(* Logix 5000 project; controller MECO9497 vendor 1 type 14 code 106 rev 21.11; software revision 21.00; part 2 of 4 *)
(* tags used below, declared in another part *)
   AAH_200 : BOOL;
   AAH_200_DELAY : TIMER;
   AAH_200_SP : REAL;
   ACKNOWLEDGE : BOOL;
   ALARM_ACK_OIT : BOOL;
   ALARM_RESET_OIT : BOOL;
   ALERT_ALARM_SU_DELAY : TIMER;
   AT_200_EU : REAL;
   COMP_AMP_ALRM_DELAY_TMR : TIMER;
   COMPRESSOR_START_CMD : BOOL;
   D_V_REMOTE_START : BOOL;
   DIST_COND_ALRM_STARTUP_TMR : TIMER;
   DSTLT_STORAGE_ENABLE_MAP : BOOL;
   DSTLT_STORAGE_ENABLE_OIT : BOOL;
   DSTLT_TEMP_ALRM_SU_DELAY : TIMER;
   E_Stop : ALIAS FOR Local:1:I.Data.0;
   E_Stop_DI_MAP : BOOL;
   ENGINEER : BOOL;
   EVAP_PRESS_CV_LIMIT : BOOL;
   EVAP_PRESS_CV_PERMISSIVE : REAL;
   EVAP_PRESS_RAMP_ONE_SHOT : BOOL;
   EVAP_PRESS_RAMP_TIMER : TIMER;
   EVAP_PRESSURE_CV_PERM : BOOL;
   EVAP_RAMP_COMPLETE : BOOL;
   EVAP_RAMP_ENABLE_DELAY_TIMER : TIMER;
   FEED_LVL_CV_LIMIT : BOOL;
   FEED_LVL_CV_LIMIT_SHUTDOWN : BOOL;
   FEED_LVL_CV_LIMIT_SHUTDOWN_DELAY : TIMER;
   FEED_LVL_CV_LIMIT_SHUTDOWN_LATCH : BOOL;
   FEED_LVL_ONE_SHOT : BOOL;
   FEED_TEM_SD_LATCH : BOOL;
   FEED_TEM_SD_TIMER : TIMER;
   FEED_TEMP_SD_ONS : BOOL;
   FEED_TEMP_STEP_DELAY : TIMER;
   HOT_STANDBY : BOOL;
   IAL_100 : BOOL;
   IAL_100_CTR : COUNTER;
   IAL_100_DELAY : TIMER;
   IAL_100_SP : REAL;
   INITIAL_SCAN_SYS_RESET : BOOL;
   INITIAL_START_STEAM_LIMIT_TMR : TIMER;
   IY_100_EU : REAL;
   LAAH_100 : BOOL;
   LAAH_100_DELAY : TIMER;
   LAAH_100_SP : DINT;
   LAAL_100 : BOOL;
   LAAL_100_DELAY : TIMER;
   LAAL_100_SP : DINT;
   LAH_100 : BOOL;
   LAH_100_AUX : BOOL;
   LAH_100_DELAY : TIMER;
   LAH_100_SP : REAL;
   LAL_100 : BOOL;
   LAL_100_DELAY : TIMER;
   LAL_100_SP : REAL;
   LB_OIL_LOW_PRESS_ALRM_DELAY : TIMER;
   LCV_100_INTERLOCK : BOOL;
   LIC_100 : PID;
   LIC_1000_CV1 : REAL;
   LIC_100_A_M_OIT : BOOL;
   LIC_100_CV2 : REAL;
   LIC_100_CV_H : BOOL;
   LIC_100_CV_N : BOOL;
   LIC_100_CV_OIT : REAL;
   LIC_100_FINAL_SP : REAL;
   LIC_100_FINAL_SP_EU : REAL;
   LIC_100_GAIN_H : BOOL;
   LIC_100_GAIN_N : BOOL;
   LIC_100_GAIN_OIT : REAL;
   LIC_100_RATE_H : BOOL;
   LIC_100_RATE_N : BOOL;
   LIC_100_RATE_OIT : REAL;
   LIC_100_RESET_H : BOOL;
   LIC_100_RESET_N : BOOL;
   LIC_100_RESET_OIT : REAL;
   LIC_100_SP_CONV : REAL;
   LIC_100_SP_EU : REAL;
   LIC_100_SP_H : BOOL;
   LIC_100_SP_N : BOOL;
   LIC_100_SP_OIT : REAL;
   LIC_100_STBY_SP : REAL;
   LIC_100_STBY_SP_EU : REAL;
   LIC_100_STBY_SP_H : BOOL;
   LIC_100_STBY_SP_N : BOOL;
   LIC_100_STBY_SP_OIT : REAL;
   LT_100_AI : ALIAS FOR Local:3:I.Ch3Data;
   LT_100_EU : REAL;
   LT_100_EU_SPAN : REAL;
   LT_100_EU_ZERO : REAL;
   M1_DI : ALIAS FOR Local:1:I.Data.1;
   M1_DI_MAP : BOOL;
   M2_DI : ALIAS FOR Local:1:I.Data.2;
   M2_DI_MAP : BOOL;
   M4_DI : ALIAS FOR Local:1:I.Data.4;
   M4_DI_MAP : BOOL;
   MAINTENANCE : BOOL;
   MCB : BOOL;
   OP_SWTCH_AUTO_DI : ALIAS FOR Local:1:I.Data.14;
   OP_SWTCH_AUTO_DI_MAP : BOOL;
   OP_SWTCH_MANUAL_DI : ALIAS FOR Local:1:I.Data.13;
   OP_SWTCH_MANUAL_DI_MAP : BOOL;
   OPERATOR : BOOL;
   PAAH_103 : BOOL;
   PAAH_103_DELAY : TIMER;
   PAAH_103_SP : REAL;
   PAAL_103 : BOOL;
   PAAL_103_DELAY : TIMER;
   PAAL_103_SP : REAL;
   PAH_103 : BOOL;
   PAH_103_AUX : BOOL;
   PAH_103_DELAY : TIMER;
   PAH_103_SP : REAL;
   PAL_103 : BOOL;
   PAL_103_DELAY : TIMER;
   PAL_103_SP : REAL;
   PAL_700 : BOOL;
   PAL_700_ALRM_DELAY : TIMER;
   PCV_103_INTERLOCK : BOOL;
   PIC_103 : PID;
   PIC_103_A_M_OIT : BOOL;
   PIC_103_CV_H : BOOL;
   PIC_103_CV_N : BOOL;
   PIC_103_CV_OIT : REAL;
   PIC_103_FINAL_SP : REAL;
   PIC_103_GAIN_H : BOOL;
   PIC_103_GAIN_N : BOOL;
   PIC_103_GAIN_OIT : REAL;
   PIC_103_RATE_H : BOOL;
   PIC_103_RATE_N : BOOL;
   PIC_103_RATE_OIT : REAL;
   PIC_103_RESET_H : BOOL;
   PIC_103_RESET_N : BOOL;
   PIC_103_RESET_OIT : REAL;
   PIC_103_SP_CONV : REAL;
   PIC_103_SP_EU : REAL;
   PIC_103_SP_H : BOOL;
   PIC_103_SP_N : BOOL;
   PIC_103_SP_OIT : REAL;
   PIC_103_STBY_SP : REAL;
   PIC_103_STBY_SP_EU : REAL;
   PIC_103_STBY_SP_H : BOOL;
   PIC_103_STBY_SP_N : BOOL;
   PIC_103_STBY_SP_OIT : REAL;
   PSL_700_DI : ALIAS FOR Local:1:I.Data.7;
   PT_103_AI : ALIAS FOR Local:3:I.Ch0Data;
   PT_103_EU : REAL;
   PT_103_EU_SPAN : REAL;
   PT_103_EU_ZERO : REAL;
   PT_103_HIGH : REAL;
   RESET : BOOL;
   SECURITY_ENABLED : BOOL;
   TAH_700 : BOOL;
   TAH_700_ALRM_DELAY : TIMER;
   TAL_200 : BOOL;
   TAL_200_DELAY : TIMER;
   TAL_200_SP : REAL;
   TIC_102 : PID;
   TIC_102_A_M_OIT : BOOL;
   TIC_102_CV_H : BOOL;
   TIC_102_CV_MIN_LIMIT : BOOL;
   TIC_102_CV_N : BOOL;
   TIC_102_CV_OIT : REAL;
   TIC_102_CV_SU_REM : DINT;
   TIC_102_CV_SU_TIMER : TIMER;
   TIC_102_GAIN_H : BOOL;
   TIC_102_GAIN_N : BOOL;
   TIC_102_GAIN_OIT : REAL;
   TIC_102_MINCV1 : REAL;
   TIC_102_MINCV2 : REAL;
   TIC_102_MINCV3 : REAL;
   TIC_102_RATE_H : BOOL;
   TIC_102_RATE_N : BOOL;
   TIC_102_RATE_OIT : REAL;
   TIC_102_RESET_H : BOOL;
   TIC_102_RESET_N : BOOL;
   TIC_102_RESET_OIT : REAL;
   TIC_102_SP_CONV : REAL;
   TIC_102_SP_EU : REAL;
   TIC_102_SP_H : BOOL;
   TIC_102_SP_N : BOOL;
   TIC_102_SP_OIT : REAL;
   TIC_102_START_CV_TIMER_SP_H : BOOL;
   TIC_102_START_CV_TIMER_SP_N : BOOL;
   TIC_102_START_CV_TIMER_SP_O : REAL;
   TSH_700_DI : ALIAS FOR Local:1:I.Data.8;
   TT_102_EU_SPAN : REAL;
   TT_102_EU_ZERO : REAL;
   TT_200_EU : REAL;
   UNIT_REMOTE_START_DI : ALIAS FOR Local:1:I.Data.12;
   UNIT_REMOTE_START_MAP : BOOL;
   UNIT_START_DI : ALIAS FOR Local:1:I.Data.10;
   UNIT_START_DI_MAP : BOOL;
   UNIT_STOP_DI : ALIAS FOR Local:1:I.Data.11;
   UNIT_STOP_DI_MAP : BOOL;
(* MainProgram, continued *)

ROUTINE EVAPORATOR_PRESSURE   (* ladder *)
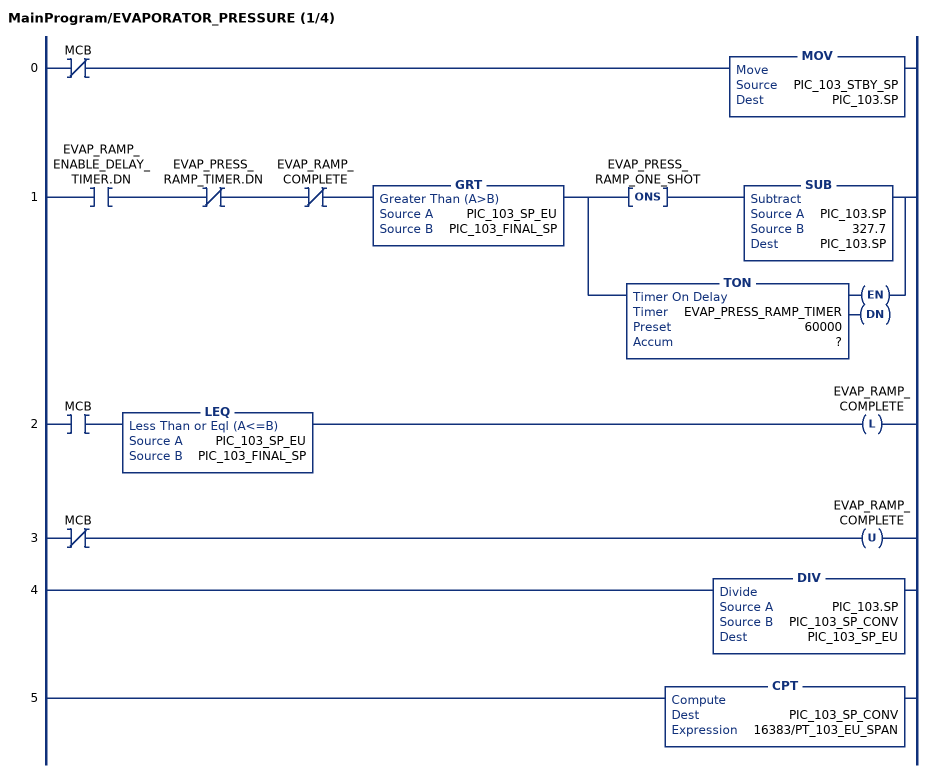
   0: XIO(MCB)MOV(PIC_103_STBY_SP,PIC_103.SP);
   1: XIC(EVAP_RAMP_ENABLE_DELAY_TIMER.DN)XIO(EVAP_PRESS_RAMP_TIMER.DN)XIO(EVAP_RAMP_COMPLETE)GRT(PIC_103_SP_EU,PIC_103_FINAL_SP)[ONS(EVAP_PRESS_RAMP_ONE_SHOT) SUB(PIC_103.SP,327.7,PIC_103.SP) ,TON(EVAP_PRESS_RAMP_TIMER,?,?) ];
   2: XIC(MCB)LEQ(PIC_103_SP_EU,PIC_103_FINAL_SP)OTL(EVAP_RAMP_COMPLETE);
   3: XIO(MCB)OTU(EVAP_RAMP_COMPLETE);
   4: DIV(PIC_103.SP,PIC_103_SP_CONV,PIC_103_SP_EU);
   5: CPT(PIC_103_SP_CONV,16383/PT_103_EU_SPAN);
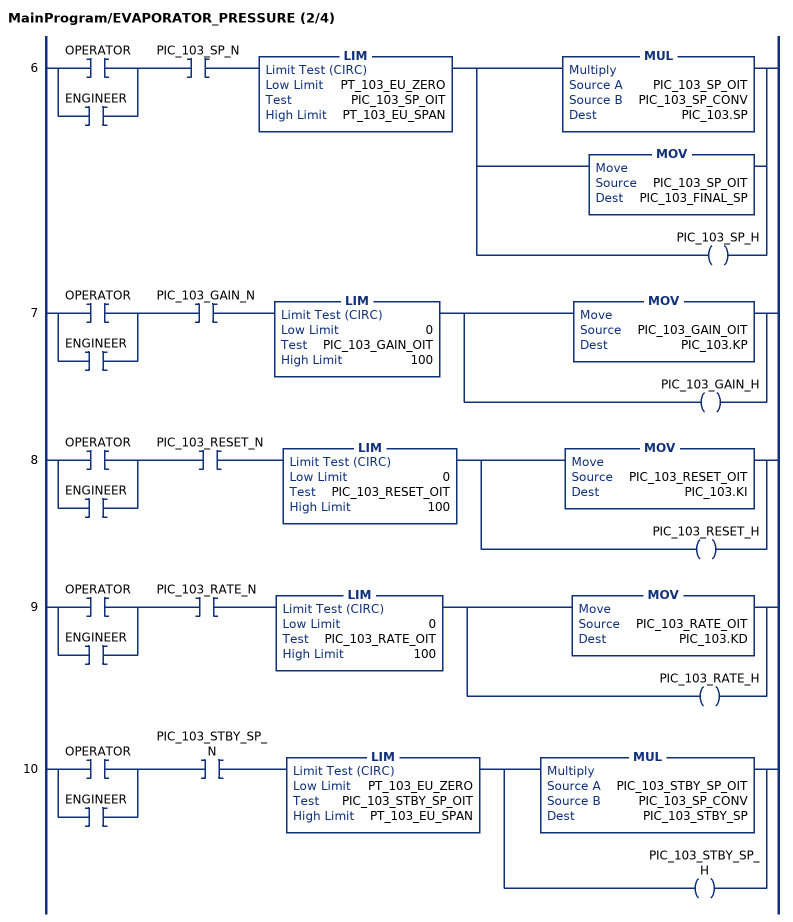
   6: [XIC(OPERATOR) ,XIC(ENGINEER) ]XIC(PIC_103_SP_N)LIM(PT_103_EU_ZERO,PIC_103_SP_OIT,PT_103_EU_SPAN)[MUL(PIC_103_SP_OIT,PIC_103_SP_CONV,PIC_103.SP) ,MOV(PIC_103_SP_OIT,PIC_103_FINAL_SP) ,OTE(PIC_103_SP_H) ];
   7: [XIC(OPERATOR) ,XIC(ENGINEER) ]XIC(PIC_103_GAIN_N)LIM(0,PIC_103_GAIN_OIT,100)[MOV(PIC_103_GAIN_OIT,PIC_103.KP) ,OTE(PIC_103_GAIN_H) ];
   8: [XIC(OPERATOR) ,XIC(ENGINEER) ]XIC(PIC_103_RESET_N)LIM(0,PIC_103_RESET_OIT,100)[MOV(PIC_103_RESET_OIT,PIC_103.KI) ,OTE(PIC_103_RESET_H) ];
   9: [XIC(OPERATOR) ,XIC(ENGINEER) ]XIC(PIC_103_RATE_N)LIM(0,PIC_103_RATE_OIT,100)[MOV(PIC_103_RATE_OIT,PIC_103.KD) ,OTE(PIC_103_RATE_H) ];
   10: [XIC(OPERATOR) ,XIC(ENGINEER) ]XIC(PIC_103_STBY_SP_N)LIM(PT_103_EU_ZERO,PIC_103_STBY_SP_OIT,PT_103_EU_SPAN)[MUL(PIC_103_STBY_SP_OIT,PIC_103_SP_CONV,PIC_103_STBY_SP) ,OTE(PIC_103_STBY_SP_H) ];
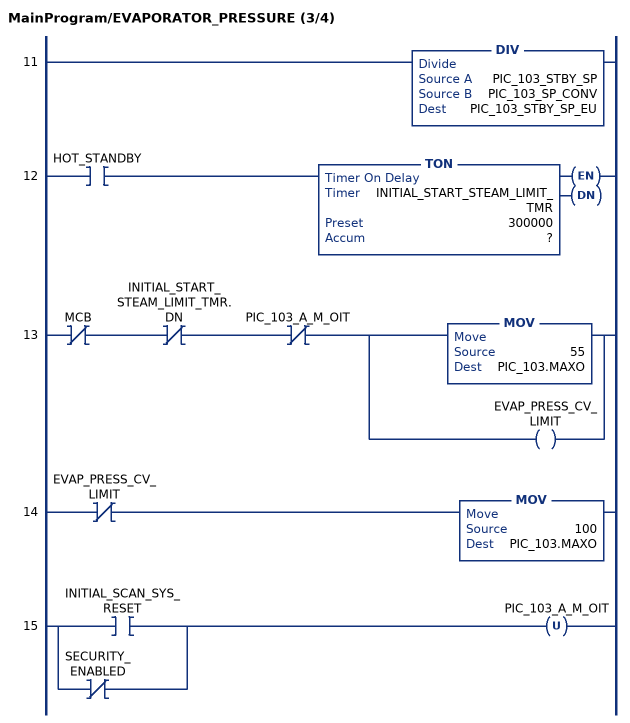
   11: DIV(PIC_103_STBY_SP,PIC_103_SP_CONV,PIC_103_STBY_SP_EU);
   12: XIC(HOT_STANDBY)TON(INITIAL_START_STEAM_LIMIT_TMR,?,?);
   13: XIO(MCB)XIO(INITIAL_START_STEAM_LIMIT_TMR.DN)XIO(PIC_103_A_M_OIT)[MOV(55,PIC_103.MAXO) ,OTE(EVAP_PRESS_CV_LIMIT) ];
   14: XIO(EVAP_PRESS_CV_LIMIT)MOV(100,PIC_103.MAXO);
   15: [XIC(INITIAL_SCAN_SYS_RESET) ,XIO(SECURITY_ENABLED) ]OTU(PIC_103_A_M_OIT);
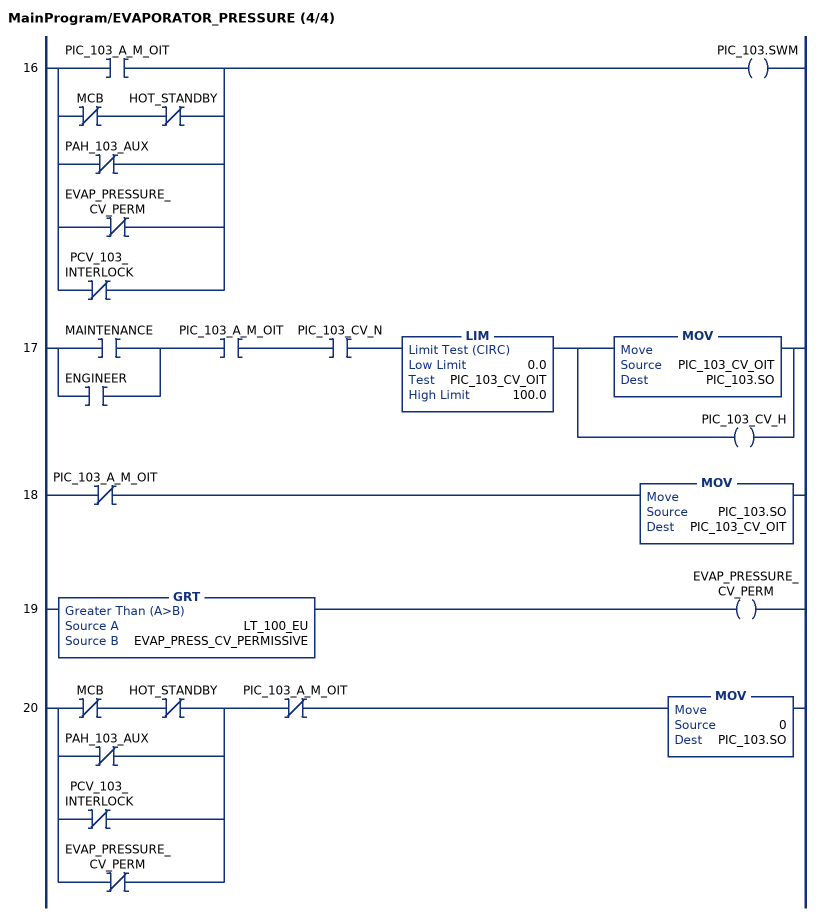
   16: [XIC(PIC_103_A_M_OIT) ,XIO(MCB) XIO(HOT_STANDBY) ,XIO(PAH_103_AUX) ,XIO(EVAP_PRESSURE_CV_PERM) ,XIO(PCV_103_INTERLOCK) ]OTE(PIC_103.SWM);
   17: [XIC(MAINTENANCE) ,XIC(ENGINEER) ]XIC(PIC_103_A_M_OIT)XIC(PIC_103_CV_N)LIM(0.0,PIC_103_CV_OIT,100.0)[MOV(PIC_103_CV_OIT,PIC_103.SO) ,OTE(PIC_103_CV_H) ];
   18: XIO(PIC_103_A_M_OIT)MOV(PIC_103.SO,PIC_103_CV_OIT);
   19: GRT(LT_100_EU,EVAP_PRESS_CV_PERMISSIVE)OTE(EVAP_PRESSURE_CV_PERM);
   20: [XIO(MCB) XIO(HOT_STANDBY) ,XIO(PAH_103_AUX) ,XIO(PCV_103_INTERLOCK) ,XIO(EVAP_PRESSURE_CV_PERM) ]XIO(PIC_103_A_M_OIT)MOV(0,PIC_103.SO);
END_ROUTINE

ROUTINE FEED_LEVEL   (* ladder *)
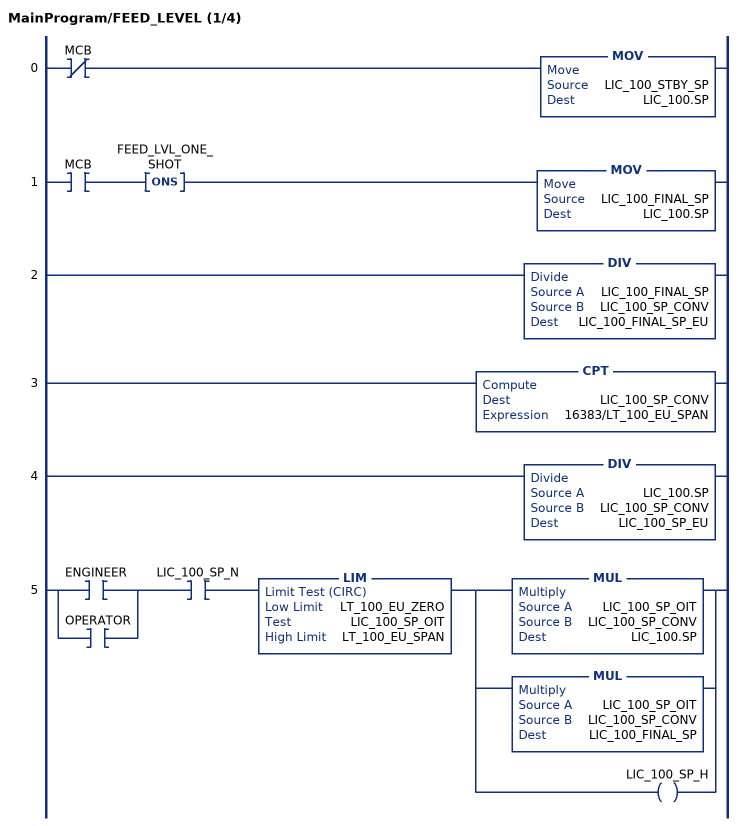
   0: XIO(MCB)MOV(LIC_100_STBY_SP,LIC_100.SP);
   1: XIC(MCB)ONS(FEED_LVL_ONE_SHOT)MOV(LIC_100_FINAL_SP,LIC_100.SP);
   2: DIV(LIC_100_FINAL_SP,LIC_100_SP_CONV,LIC_100_FINAL_SP_EU);
   3: CPT(LIC_100_SP_CONV,16383/LT_100_EU_SPAN);
   4: DIV(LIC_100.SP,LIC_100_SP_CONV,LIC_100_SP_EU);
   5: [XIC(ENGINEER) ,XIC(OPERATOR) ]XIC(LIC_100_SP_N)LIM(LT_100_EU_ZERO,LIC_100_SP_OIT,LT_100_EU_SPAN)[[MUL(LIC_100_SP_OIT,LIC_100_SP_CONV,LIC_100.SP) ,MUL(LIC_100_SP_OIT,LIC_100_SP_CONV,LIC_100_FINAL_SP) ] ,OTE(LIC_100_SP_H) ];
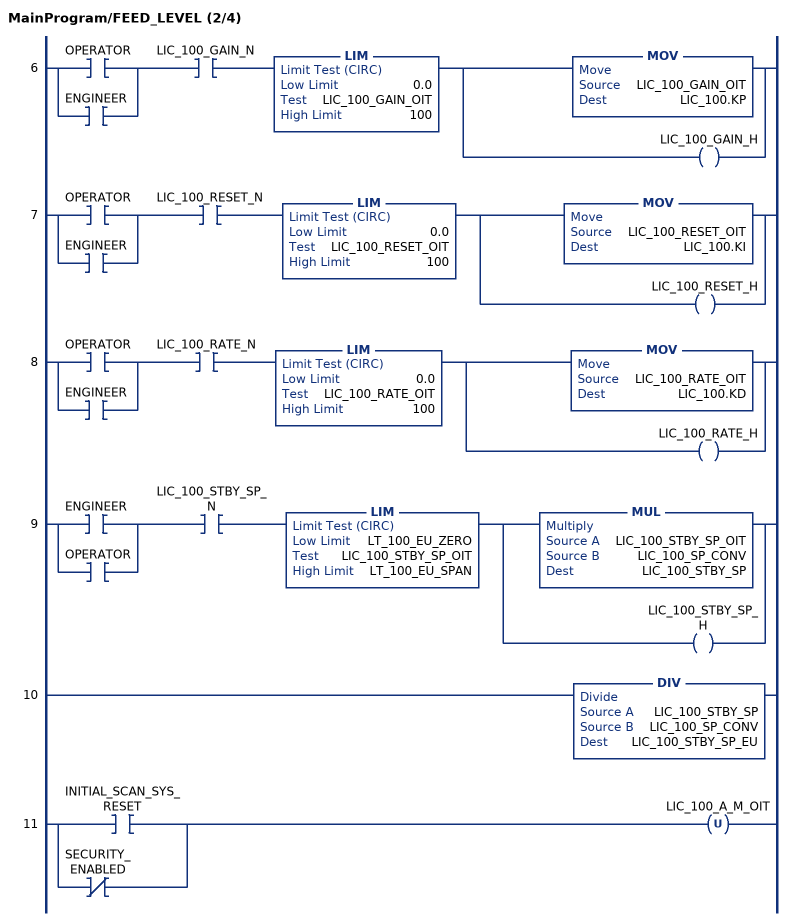
   6: [XIC(OPERATOR) ,XIC(ENGINEER) ]XIC(LIC_100_GAIN_N)LIM(0.0,LIC_100_GAIN_OIT,100)[MOV(LIC_100_GAIN_OIT,LIC_100.KP) ,OTE(LIC_100_GAIN_H) ];
   7: [XIC(OPERATOR) ,XIC(ENGINEER) ]XIC(LIC_100_RESET_N)LIM(0.0,LIC_100_RESET_OIT,100)[MOV(LIC_100_RESET_OIT,LIC_100.KI) ,OTE(LIC_100_RESET_H) ];
   8: [XIC(OPERATOR) ,XIC(ENGINEER) ]XIC(LIC_100_RATE_N)LIM(0.0,LIC_100_RATE_OIT,100)[MOV(LIC_100_RATE_OIT,LIC_100.KD) ,OTE(LIC_100_RATE_H) ];
   9: [XIC(ENGINEER) ,XIC(OPERATOR) ]XIC(LIC_100_STBY_SP_N)LIM(LT_100_EU_ZERO,LIC_100_STBY_SP_OIT,LT_100_EU_SPAN)[MUL(LIC_100_STBY_SP_OIT,LIC_100_SP_CONV,LIC_100_STBY_SP) ,OTE(LIC_100_STBY_SP_H) ];
   10: DIV(LIC_100_STBY_SP,LIC_100_SP_CONV,LIC_100_STBY_SP_EU);
   11: [XIC(INITIAL_SCAN_SYS_RESET) ,XIO(SECURITY_ENABLED) ]OTU(LIC_100_A_M_OIT);
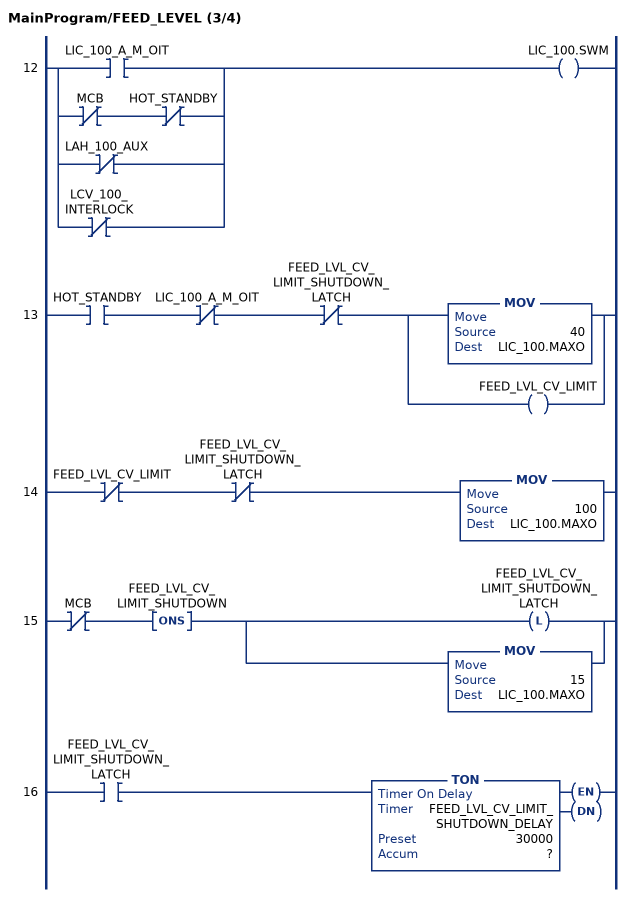
   12: [XIC(LIC_100_A_M_OIT) ,XIO(MCB) XIO(HOT_STANDBY) ,XIO(LAH_100_AUX) ,XIO(LCV_100_INTERLOCK) ]OTE(LIC_100.SWM);
   13: XIC(HOT_STANDBY)XIO(LIC_100_A_M_OIT)XIO(FEED_LVL_CV_LIMIT_SHUTDOWN_LATCH)[MOV(40,LIC_100.MAXO) ,OTE(FEED_LVL_CV_LIMIT) ];
   14: XIO(FEED_LVL_CV_LIMIT)XIO(FEED_LVL_CV_LIMIT_SHUTDOWN_LATCH)MOV(100,LIC_100.MAXO);
   15: XIO(MCB)ONS(FEED_LVL_CV_LIMIT_SHUTDOWN)[OTL(FEED_LVL_CV_LIMIT_SHUTDOWN_LATCH) ,MOV(15,LIC_100.MAXO) ];
   16: XIC(FEED_LVL_CV_LIMIT_SHUTDOWN_LATCH)TON(FEED_LVL_CV_LIMIT_SHUTDOWN_DELAY,?,?);
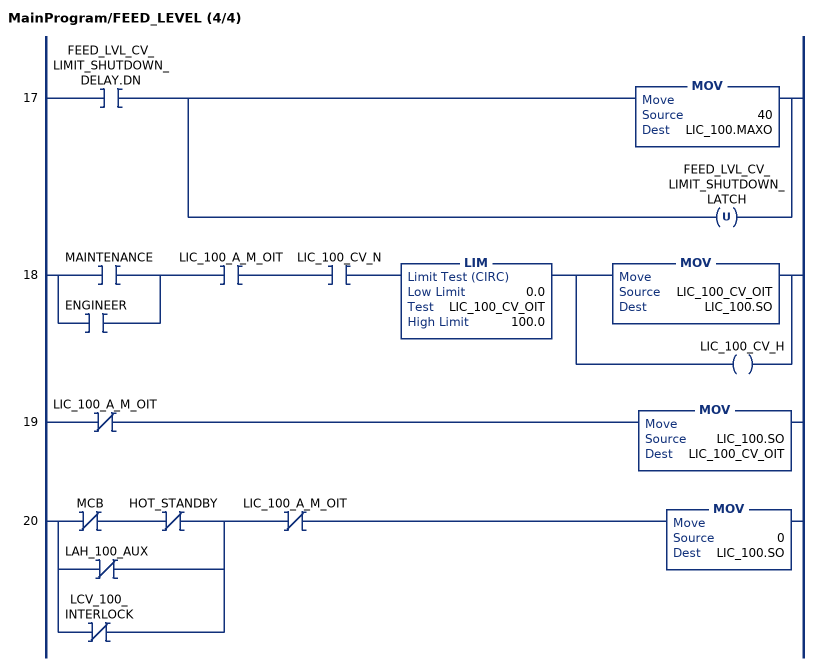
   17: XIC(FEED_LVL_CV_LIMIT_SHUTDOWN_DELAY.DN)[MOV(40,LIC_100.MAXO) ,OTU(FEED_LVL_CV_LIMIT_SHUTDOWN_LATCH) ];
   18: [XIC(MAINTENANCE) ,XIC(ENGINEER) ]XIC(LIC_100_A_M_OIT)XIC(LIC_100_CV_N)LIM(0.0,LIC_100_CV_OIT,100.0)[MOV(LIC_100_CV_OIT,LIC_100.SO) ,OTE(LIC_100_CV_H) ];
   19: XIO(LIC_100_A_M_OIT)MOV(LIC_100.SO,LIC_100_CV_OIT);
   20: [XIO(MCB) XIO(HOT_STANDBY) ,XIO(LAH_100_AUX) ,XIO(LCV_100_INTERLOCK) ]XIO(LIC_100_A_M_OIT)MOV(0,LIC_100.SO);
END_ROUTINE

ROUTINE FEED_TEMPERATURE   (* ladder *)
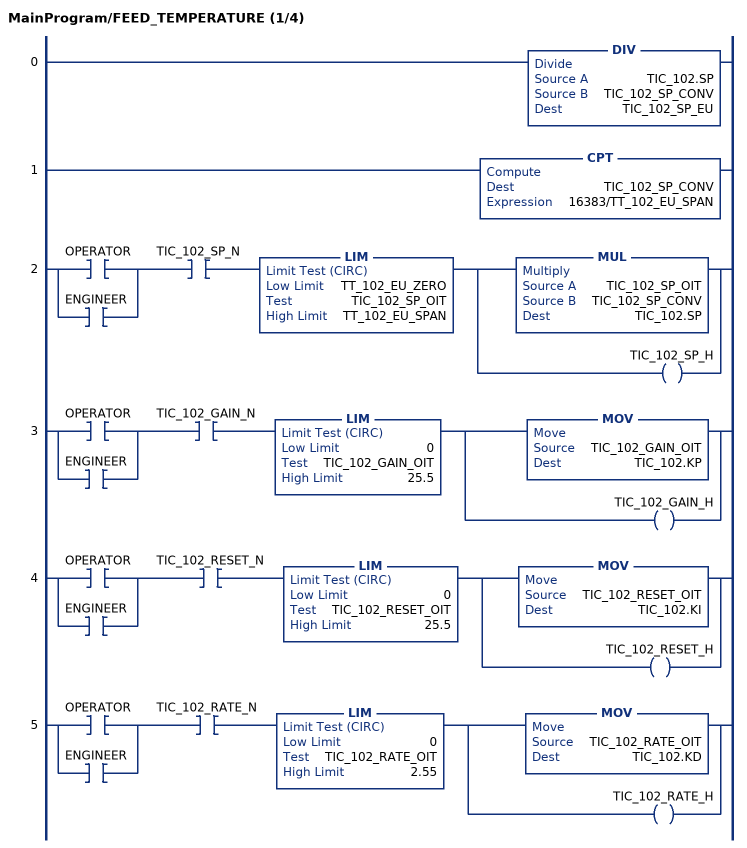
   0: DIV(TIC_102.SP,TIC_102_SP_CONV,TIC_102_SP_EU);
   1: CPT(TIC_102_SP_CONV,16383/TT_102_EU_SPAN);
   2: [XIC(OPERATOR) ,XIC(ENGINEER) ]XIC(TIC_102_SP_N)LIM(TT_102_EU_ZERO,TIC_102_SP_OIT,TT_102_EU_SPAN)[MUL(TIC_102_SP_OIT,TIC_102_SP_CONV,TIC_102.SP) ,OTE(TIC_102_SP_H) ];
   3: [XIC(OPERATOR) ,XIC(ENGINEER) ]XIC(TIC_102_GAIN_N)LIM(0,TIC_102_GAIN_OIT,25.5)[MOV(TIC_102_GAIN_OIT,TIC_102.KP) ,OTE(TIC_102_GAIN_H) ];
   4: [XIC(OPERATOR) ,XIC(ENGINEER) ]XIC(TIC_102_RESET_N)LIM(0,TIC_102_RESET_OIT,25.5)[MOV(TIC_102_RESET_OIT,TIC_102.KI) ,OTE(TIC_102_RESET_H) ];
   5: [XIC(OPERATOR) ,XIC(ENGINEER) ]XIC(TIC_102_RATE_N)LIM(0,TIC_102_RATE_OIT,2.55)[MOV(TIC_102_RATE_OIT,TIC_102.KD) ,OTE(TIC_102_RATE_H) ];
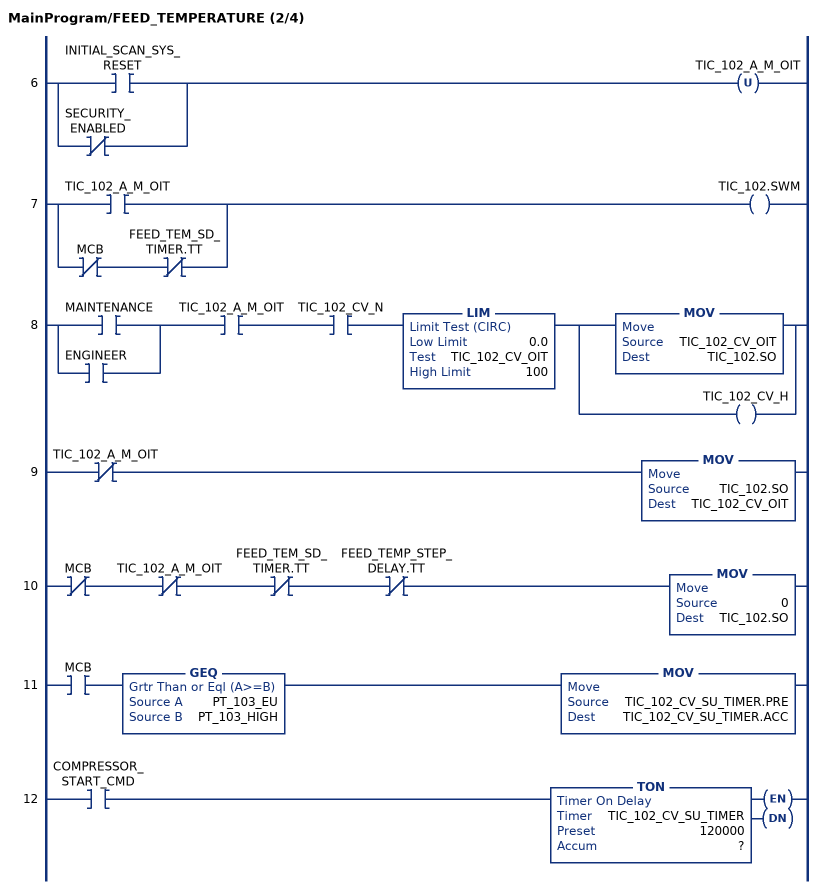
   6: [XIC(INITIAL_SCAN_SYS_RESET) ,XIO(SECURITY_ENABLED) ]OTU(TIC_102_A_M_OIT);
   7: [XIC(TIC_102_A_M_OIT) ,XIO(MCB) XIO(FEED_TEM_SD_TIMER.TT) ]OTE(TIC_102.SWM);
   8: [XIC(MAINTENANCE) ,XIC(ENGINEER) ]XIC(TIC_102_A_M_OIT)XIC(TIC_102_CV_N)LIM(0.0,TIC_102_CV_OIT,100)[MOV(TIC_102_CV_OIT,TIC_102.SO) ,OTE(TIC_102_CV_H) ];
   9: XIO(TIC_102_A_M_OIT)MOV(TIC_102.SO,TIC_102_CV_OIT);
   10: XIO(MCB)XIO(TIC_102_A_M_OIT)XIO(FEED_TEM_SD_TIMER.TT)XIO(FEED_TEMP_STEP_DELAY.TT)MOV(0,TIC_102.SO);
   11: XIC(MCB)GEQ(PT_103_EU,PT_103_HIGH)MOV(TIC_102_CV_SU_TIMER.PRE,TIC_102_CV_SU_TIMER.ACC);
   12: XIC(COMPRESSOR_START_CMD)TON(TIC_102_CV_SU_TIMER,?,?);
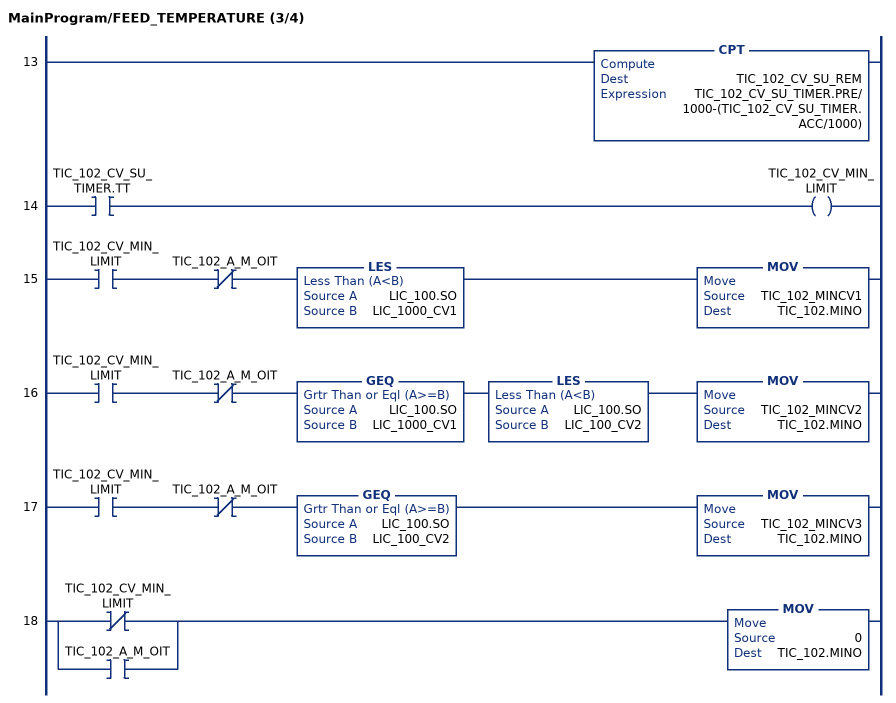
   13: CPT(TIC_102_CV_SU_REM,TIC_102_CV_SU_TIMER.PRE/1000-(TIC_102_CV_SU_TIMER.ACC/1000));
   14: XIC(TIC_102_CV_SU_TIMER.TT)OTE(TIC_102_CV_MIN_LIMIT);
   15: XIC(TIC_102_CV_MIN_LIMIT)XIO(TIC_102_A_M_OIT)LES(LIC_100.SO,LIC_1000_CV1)MOV(TIC_102_MINCV1,TIC_102.MINO);
   16: XIC(TIC_102_CV_MIN_LIMIT)XIO(TIC_102_A_M_OIT)GEQ(LIC_100.SO,LIC_1000_CV1)LES(LIC_100.SO,LIC_100_CV2)MOV(TIC_102_MINCV2,TIC_102.MINO);
   17: XIC(TIC_102_CV_MIN_LIMIT)XIO(TIC_102_A_M_OIT)GEQ(LIC_100.SO,LIC_100_CV2)MOV(TIC_102_MINCV3,TIC_102.MINO);
   18: [XIO(TIC_102_CV_MIN_LIMIT) ,XIC(TIC_102_A_M_OIT) ]MOV(0,TIC_102.MINO);
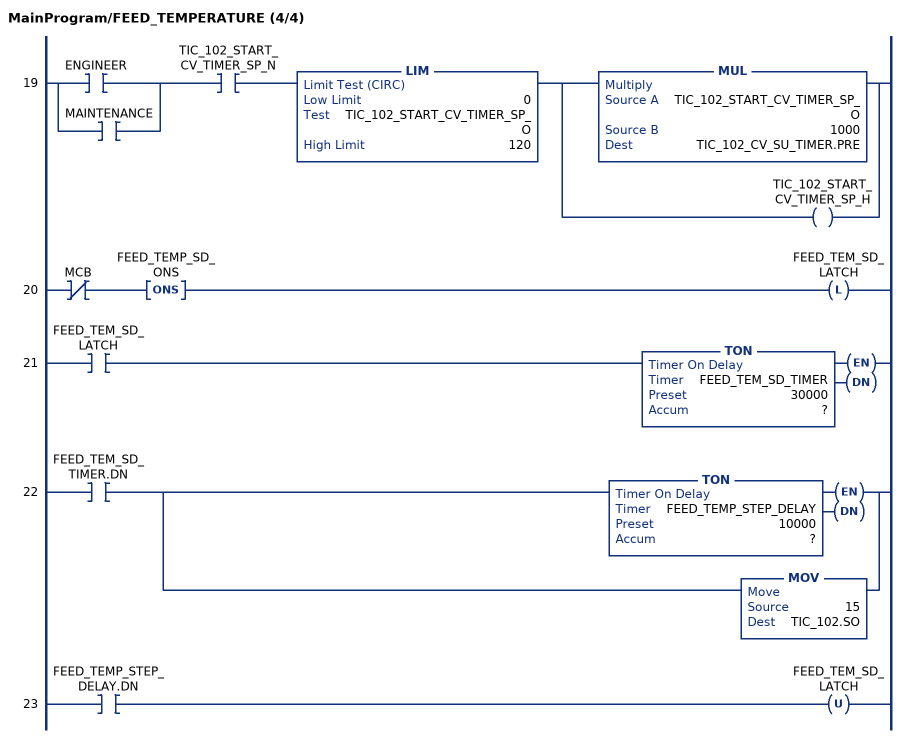
   19: [XIC(ENGINEER) ,XIC(MAINTENANCE) ]XIC(TIC_102_START_CV_TIMER_SP_N)LIM(0,TIC_102_START_CV_TIMER_SP_O,120)[MUL(TIC_102_START_CV_TIMER_SP_O,1000,TIC_102_CV_SU_TIMER.PRE) ,OTE(TIC_102_START_CV_TIMER_SP_H) ];
   20: XIO(MCB)ONS(FEED_TEMP_SD_ONS)OTL(FEED_TEM_SD_LATCH);
   21: XIC(FEED_TEM_SD_LATCH)TON(FEED_TEM_SD_TIMER,?,?);
   22: XIC(FEED_TEM_SD_TIMER.DN)[TON(FEED_TEMP_STEP_DELAY,?,?) ,MOV(15,TIC_102.SO) ];
   23: XIC(FEED_TEMP_STEP_DELAY.DN)OTU(FEED_TEM_SD_LATCH);
END_ROUTINE

ROUTINE INPUT_MAP   (* ladder *)
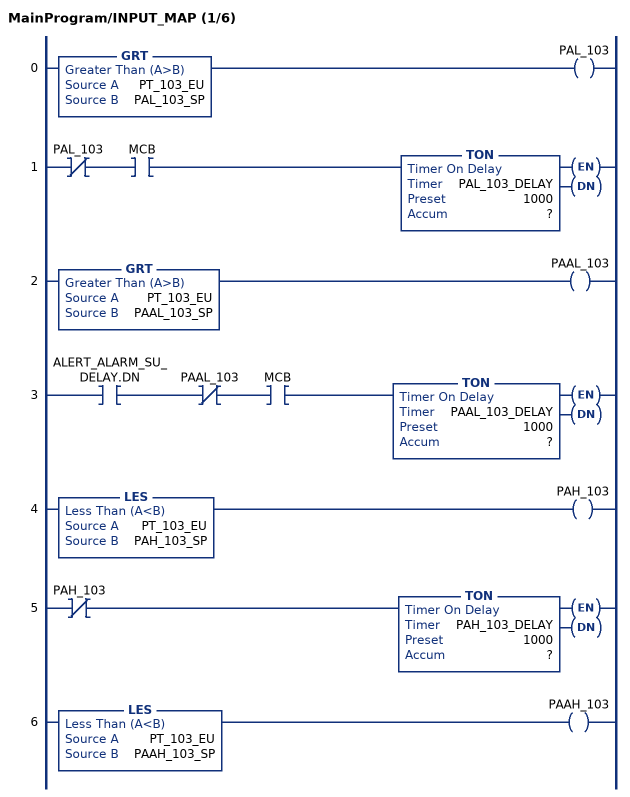
   0: GRT(PT_103_EU,PAL_103_SP)OTE(PAL_103);
   1: XIO(PAL_103)XIC(MCB)TON(PAL_103_DELAY,?,?);
   2: GRT(PT_103_EU,PAAL_103_SP)OTE(PAAL_103);
   3: XIC(ALERT_ALARM_SU_DELAY.DN)XIO(PAAL_103)XIC(MCB)TON(PAAL_103_DELAY,?,?);
   4: LES(PT_103_EU,PAH_103_SP)OTE(PAH_103);
   5: XIO(PAH_103)TON(PAH_103_DELAY,?,?);
   6: LES(PT_103_EU,PAAH_103_SP)OTE(PAAH_103);
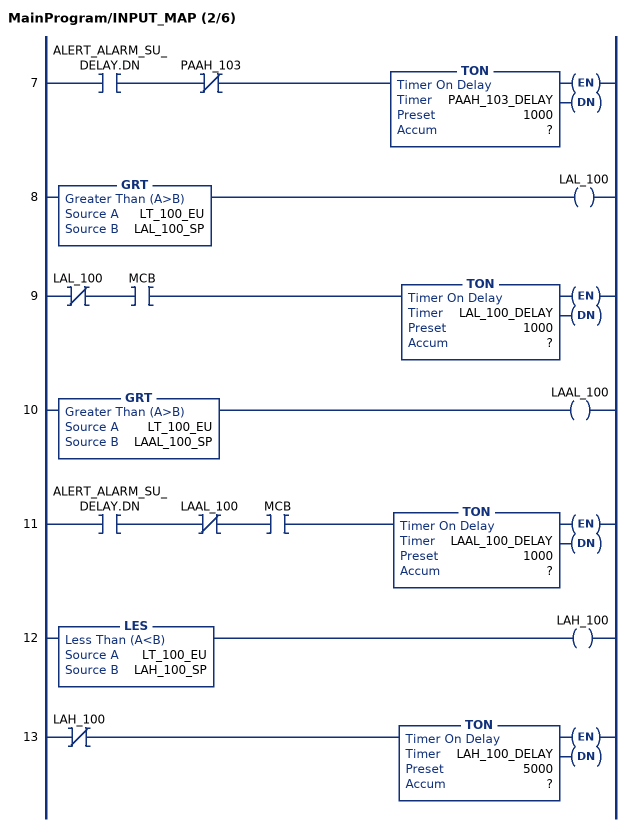
   7: XIC(ALERT_ALARM_SU_DELAY.DN)XIO(PAAH_103)TON(PAAH_103_DELAY,?,?);
   8: GRT(LT_100_EU,LAL_100_SP)OTE(LAL_100);
   9: XIO(LAL_100)XIC(MCB)TON(LAL_100_DELAY,?,?);
   10: GRT(LT_100_EU,LAAL_100_SP)OTE(LAAL_100);
   11: XIC(ALERT_ALARM_SU_DELAY.DN)XIO(LAAL_100)XIC(MCB)TON(LAAL_100_DELAY,?,?);
   12: LES(LT_100_EU,LAH_100_SP)OTE(LAH_100);
   13: XIO(LAH_100)TON(LAH_100_DELAY,?,?);
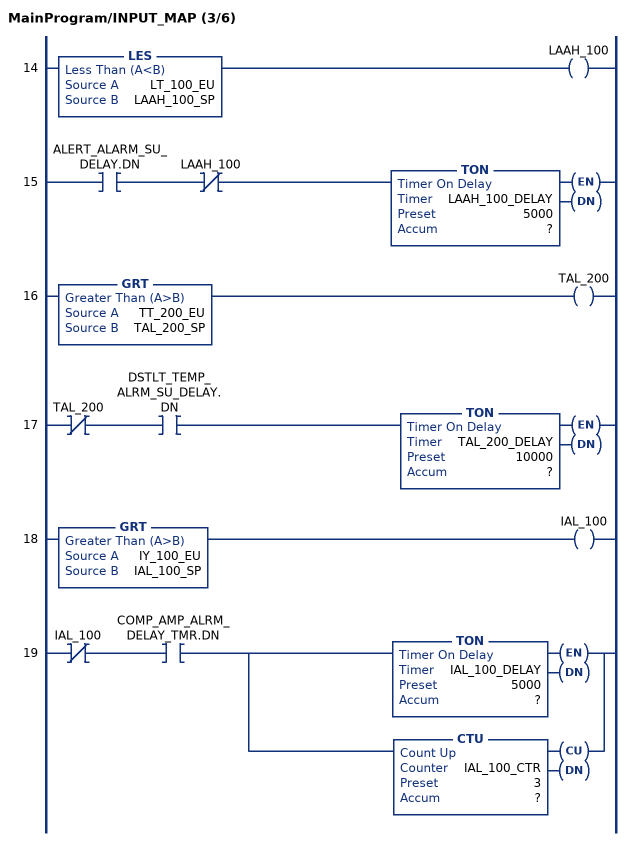
   14: LES(LT_100_EU,LAAH_100_SP)OTE(LAAH_100);
   15: XIC(ALERT_ALARM_SU_DELAY.DN)XIO(LAAH_100)TON(LAAH_100_DELAY,?,?);
   16: GRT(TT_200_EU,TAL_200_SP)OTE(TAL_200);
   17: XIO(TAL_200)XIC(DSTLT_TEMP_ALRM_SU_DELAY.DN)TON(TAL_200_DELAY,?,?);
   18: GRT(IY_100_EU,IAL_100_SP)OTE(IAL_100);
   19: XIO(IAL_100)XIC(COMP_AMP_ALRM_DELAY_TMR.DN)[TON(IAL_100_DELAY,?,?) ,CTU(IAL_100_CTR,?,?) ];
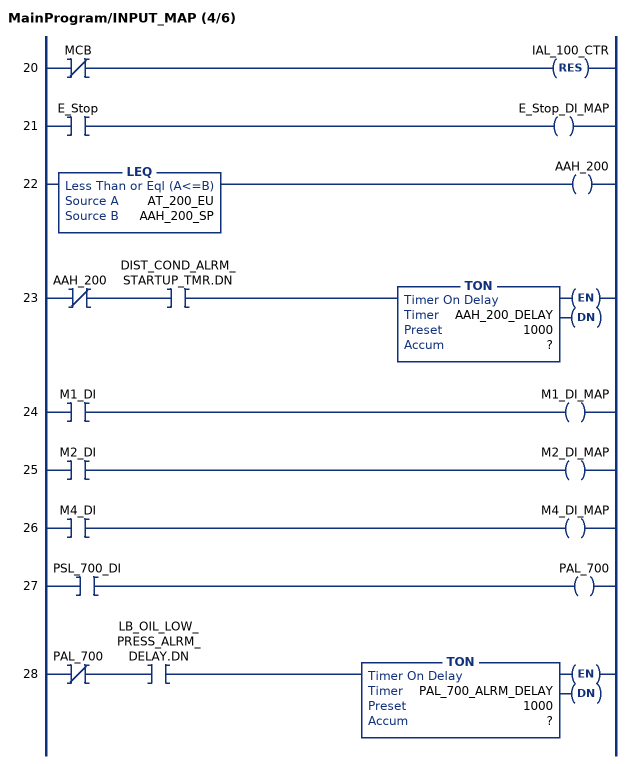
   20: XIO(MCB)RES(IAL_100_CTR);
   21: XIC(E_Stop)OTE(E_Stop_DI_MAP);
   22: LEQ(AT_200_EU,AAH_200_SP)OTE(AAH_200);
   23: XIO(AAH_200)XIC(DIST_COND_ALRM_STARTUP_TMR.DN)TON(AAH_200_DELAY,?,?);
   24: XIC(M1_DI)OTE(M1_DI_MAP);
   25: XIC(M2_DI)OTE(M2_DI_MAP);
   26: XIC(M4_DI)OTE(M4_DI_MAP);
   27: XIC(PSL_700_DI)OTE(PAL_700);
   28: XIO(PAL_700)XIC(LB_OIL_LOW_PRESS_ALRM_DELAY.DN)TON(PAL_700_ALRM_DELAY,?,?);
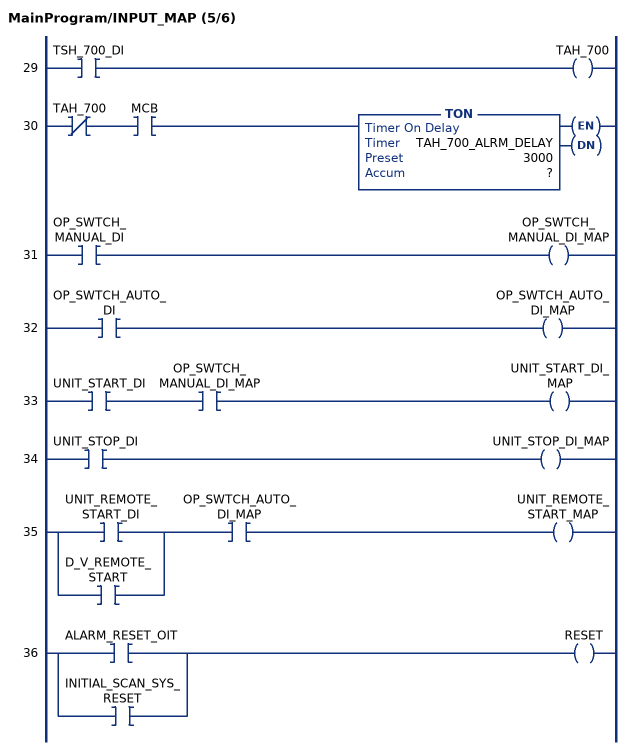
   29: XIC(TSH_700_DI)OTE(TAH_700);
   30: XIO(TAH_700)XIC(MCB)TON(TAH_700_ALRM_DELAY,?,?);
   31: XIC(OP_SWTCH_MANUAL_DI)OTE(OP_SWTCH_MANUAL_DI_MAP);
   32: XIC(OP_SWTCH_AUTO_DI)OTE(OP_SWTCH_AUTO_DI_MAP);
   33: XIC(UNIT_START_DI)XIC(OP_SWTCH_MANUAL_DI_MAP)OTE(UNIT_START_DI_MAP);
   34: XIC(UNIT_STOP_DI)OTE(UNIT_STOP_DI_MAP);
   35: [XIC(UNIT_REMOTE_START_DI) ,XIC(D_V_REMOTE_START) ]XIC(OP_SWTCH_AUTO_DI_MAP)OTE(UNIT_REMOTE_START_MAP);
   36: [XIC(ALARM_RESET_OIT) ,XIC(INITIAL_SCAN_SYS_RESET) ]OTE(RESET);
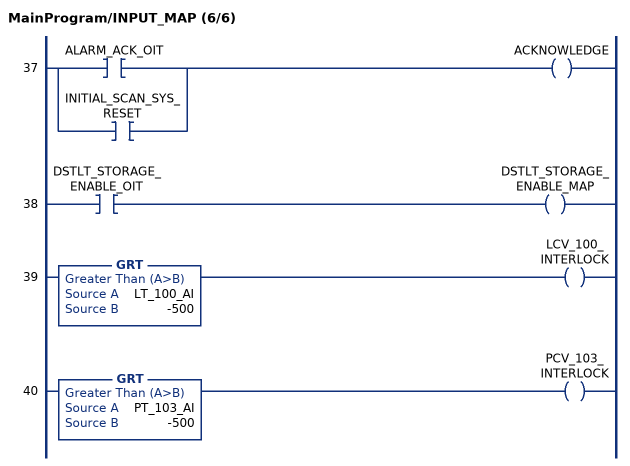
   37: [XIC(ALARM_ACK_OIT) ,XIC(INITIAL_SCAN_SYS_RESET) ]OTE(ACKNOWLEDGE);
   38: XIC(DSTLT_STORAGE_ENABLE_OIT)OTE(DSTLT_STORAGE_ENABLE_MAP);
   39: GRT(LT_100_AI,-500)OTE(LCV_100_INTERLOCK);
   40: GRT(PT_103_AI,-500)OTE(PCV_103_INTERLOCK);
END_ROUTINE
